(* IEC 61131-3 sources: s7-to-codesys/src/POUs/S7Compat/F_S5CounterBin, 1 file *)

(* ---- F_S5CounterBin.decl.st ---- *)
// Назначение: L C n — значение счётчика S5 двоичным числом (0…999).
// Автор:      kr0nsch
// Версия:     1.2.0
// Документ:   docs/MAPPING_STL.md, правило s5.counter
FUNCTION F_S5CounterBin : WORD
VAR_INPUT
    stCounter : ST_S5Counter;   // счётчик (GVL_S5Counters.aCounter[n])
END_VAR
